// TIA Portal V18 export
DATA_BLOCK "VERIFICA INTERLOCK"   // DB200
{ S7_Optimized_Access := 'TRUE' }
// stored: MemoryReserve 100
   VAR
      INTERLOCK : Array[0..10] of Struct
         STATION : Int;
         EQUIPAMENTO : Int;
         SINAL : Int;
      END_STRUCT;
      "ATIVA FOR" : Bool;
      modezone : Int;
   END_VAR
BEGIN
END_DATA_BLOCK
